Fanuc KAREL source: ko00108.compact.KL

PROGRAM KO00108
%STACKSIZE=65535
%PRIORITY=65535
%NOLOCKGROUP
VAR
A : REAL
B : REAL
OUT : REAL
BEGIN
A=1
B=2
OUT=ATAN2(A,B)
END KO00108
